(* IEC 61131-3 sources: rusty/tests/integration/data/json, 3 files *)

(* ---- program_with_expressions.st ---- *)
PROGRAM name
(1 + 2) * (3 + 4);
END_PROGRAM

(* ---- program_with_variables.st ---- *)
PROGRAM hello
VAR
   x : INT;
   y : BOOL;
END_VAR
   IF x = 2 THEN
      x := 3;
   END_IF
END_PROGRAM

(* ---- simple_program.st ---- *)
PROGRAM prg
    VAR
        a : INT;
        b : REAL;
    END_VAR
    b := 1.5;
    a := INT#b;
END_PROGRAM
